Fanuc KAREL source: kb00007.KL

-- PROVISIONAL review KL for V940-1; original PC SHA256 0e8027ba97894a2228bac0daad2c75cc7f2703da801fc14289a9be554f262da2
-- Incomplete behavior may be omitted. Consult companion uncertainty JSON. Do not deploy.
PROGRAM KB00007
%NOLOCKGROUP
BEGIN
  -- V9_ZERO_TABLE_METADATA_HINT layout=0002_ascii; no indexed target words; source/name/runtime held
  -- UNRESOLVED_PC offsets 5-28; opcodes 27,22,1C,31,4A
  -- UNRESOLVED_PC offsets 33-37; opcodes 7F
END KB00007
